Fanuc KAREL source: ko00069.KL

-- PROVISIONAL review KL for V770-1; original PC SHA256 965c70ec17ae93b2553be2dbd9bf998d5721ce7db8dd7123341ec2a7853e820c
-- Incomplete behavior may be omitted. Consult companion uncertainty JSON. Do not deploy.
PROGRAM KO00069
%NOLOCKGROUP
BEGIN
  -- UNRESOLVED_PC offsets 5-12; opcodes 9D,23
  -- UNRESOLVED_PC offsets 17-66; opcodes 27,22,1C,27,49,7E,AD,22,31,7E,4A
  -- UNRESOLVED_PC offsets 71-75; opcodes 7F
END KO00069
